Fanuc KAREL source: kd00073.KL

-- PROVISIONAL review KL for V1013-1; original PC SHA256 461de030c76bfdc21287e07158c3bff1c9f8414620ad55adfb88fa4050f9353f
-- Incomplete behavior may be omitted. Consult companion uncertainty JSON. Do not deploy.
PROGRAM KD00073
%NOLOCKGROUP
VAR
  I : INTEGER
  J : INTEGER
  B : BOOLEAN
  R : REAL
  S : STRING[80]
BEGIN
  -- UNRESOLVED_PC offsets 5-12; opcodes 9C,23
  -- UNRESOLVED_PC offsets 22-36; opcodes 21,9D,52,23
  -- UNRESOLVED_PC offsets 41-58; opcodes 21,2E,5B,79
  -- UNRESOLVED_PC offsets 63-67; opcodes 7F
END KD00073
